Fanuc KAREL source: kb00114.KL

PROGRAM KB00114
%STACKSIZE=65535
%PRIORITY=65535
%NOLOCKGROUP
VAR
P1 : STRING[80]
P2 : INTEGER
BEGIN
P1='A'
P2=1
KCL_NO_WAIT(P1,P2)
END KB00114
